FUNCTION_BLOCK TableRotateQI (* Composite Function Block Type *)
  (* Standard: 61499-2 *)
  (* Version 0.0, 7/2/2026, template *)
  PACKAGE Main;
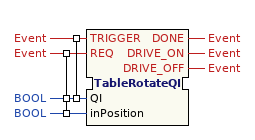
  EVENT_INPUT
    TRIGGER WITH QI; (* Initialization Request *)
    REQ WITH QI, inPosition; (* Normal Execution Request *)
  END_EVENT
  EVENT_OUTPUT
    DONE; (* Initialization Confirm *)
    DRIVE_ON; (* Execution Confirmation *)
    DRIVE_OFF;
  END_EVENT
  VAR_INPUT
    QI : BOOL; (* Input event qualifier *)
    inPosition : BOOL;
  END_VAR
  FBS
    FB1 : TableRotate;
    FB2 : E_DELAY(DT := T#500ms);
    FB3 : E_SWITCH;
  END_FBS
  EVENT_CONNECTIONS
    FB1.54922CD39726F432 TO DRIVE_ON;
    FB1.20E8908D046FFBAB TO DRIVE_OFF;
    FB1.B42838BDBF746833 TO FB2.START;
    FB3.EO0 TO FB1.3EB595A19E7C967B;
    FB3.EO1 TO DONE;
    REQ TO FB1.55C5B35594136179;
    TRIGGER TO FB1.3EB595A19E7C967B;
    FB2.EO TO FB3.EI;
  END_CONNECTIONS
  DATA_CONNECTIONS
    QI TO FB3.G;
    inPosition TO FB1.3EAF9B6241519430;
  END_CONNECTIONS
END_FUNCTION_BLOCK
